(* IEC 61131-3 sources: PLC-Static-Analysis/modules/plc-rules/src/test/resources/PLCA-L011, 2 files *)

(* ---- compliant.st ---- *)
PROGRAM P_L011ok
VAR
    n : INT;
    m : INT;
    r : REAL;
    b : BOOL;
    c : BOOL;
    q : BOOL;
END_VAR
IF n < 100 THEN
    q := TRUE;
ELSIF n >= 100 THEN
    q := FALSE;
END_IF
IF n < 0 THEN
    q := TRUE;
ELSIF n > 10 THEN
    q := FALSE;
END_IF
IF n < 0 THEN
    q := TRUE;
ELSIF n > 0 THEN
    q := FALSE;
ELSE
    b := TRUE;
END_IF
IF n <> 0 THEN
    IF n < 0 THEN
        q := TRUE;
    ELSIF n > 0 THEN
        q := FALSE;
    END_IF
END_IF
IF n = 1 THEN
    q := TRUE;
ELSIF n = 2 THEN
    q := FALSE;
END_IF
END_PROGRAM

(* ---- noncompliant.st ---- *)
PROGRAM P_L011
VAR
    n : INT;
    m : INT;
    r : REAL;
    b : BOOL;
    c : BOOL;
    q : BOOL;
END_VAR
IF n < 100 THEN // PLCA-L011
    q := TRUE;
ELSIF n > 100 THEN
    q := FALSE;
END_IF
IF n > m THEN // PLCA-L011
    q := TRUE;
ELSIF n < m THEN
    q := FALSE;
END_IF
IF r < 0.0 THEN // PLCA-L011
    q := TRUE;
ELSIF r > 0.0 THEN
    q := FALSE;
END_IF
END_PROGRAM
